Fanuc KAREL source: KT00744.KL

PROGRAM KT00744
%NOLOCKGROUP
VAR
  ARG: ARRAY[4] OF XYZWPR
  OUT: BOOLEAN
BEGIN
  OUT = UNINIT(ARG)
END KT00744
